(* IEC 61131-3 sources: JingjiangArm/moonboxpro_arm_8.4/Application/Application/任务列表/LogTask/粗采样保存/调用功能, 2 files *)

(* ---- KS_FetchNextSampleDataPtr.st ---- *)
(*@CES
Name=KS_FetchNextSampleDataPtr
Type=FunctionBlock
TypeGuid=6f9dac99-8de1-4efc-8465-68ac443b7d08
Guid=600b6e6a-0af7-4a30-ab9c-796b863be3cd
HasDeclaration=True
HasImplementation=True
*)
{DECLARATION}
FUNCTION KS_FetchNextSampleDataPtr : BOOL
VAR_INPUT
	i_pstStSampleDataForTest: POINTER TO StSampleDataForTest;
	i_ppbyRS_T1: POINTER TO POINTER TO BYTE;(* 粗采样T1数据起点 *)
	i_ppbyRS_T2: POINTER TO POINTER TO BYTE;(* 粗采样T2数据起点 *)
	i_ppbyFS_T1: POINTER TO POINTER TO BYTE;(* 精采样T1数据起点 *)
	i_ppbyFS_T2: POINTER TO POINTER TO BYTE;(* 精采样T2数据起点 *)
END_VAR
VAR
	xResult: BOOL;
	byIDX_Tmp: BYTE;
END_VAR
{IMPLEMENTATION}
IF i_pstStSampleDataForTest<>0 AND
	i_ppbyRS_T1<>0 AND
	i_ppbyRS_T2<>0 AND
	i_ppbyFS_T1<>0 AND
	i_ppbyFS_T2<>0 THEN

	xResult:= TRUE;

	(* 将当前数据位置反馈到出口参数 *)
	byIDX_Tmp:= i_pstStSampleDataForTest^.byIdx AND 7;(* 只取低3位 *)

	(* 粗采样 *)
	i_ppbyRS_T1^:= ADR(i_pstStSampleDataForTest^.abyBuf_Rs[byIDX_Tmp,   1]);
	i_ppbyRS_T2^:= ADR(i_pstStSampleDataForTest^.abyBuf_Rs[byIDX_Tmp,4001]);

	(* 精采样 *)
	i_ppbyFS_T1^:= ADR(i_pstStSampleDataForTest^.abyBuf_Fs[byIDX_Tmp,   1]);
	i_ppbyFS_T2^:= ADR(i_pstStSampleDataForTest^.abyBuf_Fs[byIDX_Tmp,4001]);

	(* go next *)
	i_pstStSampleDataForTest^.byIdx:= i_pstStSampleDataForTest^.byIdx+1;
ELSE
	xResult:= FALSE;
END_IF
KS_FetchNextSampleDataPtr:= xResult;

(* ---- KS_MallocMemAndInstallSampleDataFromFile.st ---- *)
(*@CES
Name=KS_MallocMemAndInstallSampleDataFromFile
Type=FunctionBlock
TypeGuid=6f9dac99-8de1-4efc-8465-68ac443b7d08
Guid=69c33b95-f0e0-43d2-8407-04367f5534f4
HasDeclaration=True
HasImplementation=True
*)
{DECLARATION}
FUNCTION KS_MallocMemAndInstallSampleDataFromFile : DWORD
VAR_INPUT
	i_sFilename_Rs_demo: STRING := '\cpac\rs.demo';
	i_sFilename_Fs_demo: STRING := '\cpac\fs.demo';
END_VAR
VAR
	iN: INT;
	dwMemHdl: DWORD;(* 内存句柄 *)
	dwFileHdl: DWORD;(* 文件句柄 *)
	diSize_Rs_demo: DINT;
	diSize_Fs_demo: DINT;
	pstStSampleDataForTest: POINTER TO StSampleDataForTest := 0;
END_VAR
{IMPLEMENTATION}
dwMemHdl:= SysMemAlloc(SIZEOF(pstStSampleDataForTest^));
pstStSampleDataForTest:= dwMemHdl;
IF pstStSampleDataForTest<>0 THEN
	(* 粗采样 *)
	diSize_Rs_demo:= SysFileGetSize(i_sFilename_Rs_demo);
	IF diSize_Rs_demo=16#10000 THEN(* 文件必须64kB *)
		dwFileHdl:= SysFileOpen(i_sFilename_Rs_demo, 'r');
		IF dwFileHdl<>0 THEN
			FOR iN:=1 TO 8 BY 1 DO
				SysFileSetPos(dwFileHdl, INT_TO_DWORD(iN-1)*8192);(* T1 *)
				SysFileRead(dwFileHdl, ADR(pstStSampleDataForTest^.abyBuf_Rs[iN-1,   1]), 4000);
				SysFileSetPos(dwFileHdl, INT_TO_DWORD(iN-1)*8192+4096);(* T2 *)
				SysFileRead(dwFileHdl, ADR(pstStSampleDataForTest^.abyBuf_Rs[iN-1,4001]), 4000);
			END_FOR
			SysFileClose(dwFileHdl);
		END_IF
	END_IF

	(* 精采样 *)
	diSize_Fs_demo:= SysFileGetSize(i_sFilename_Fs_demo);
	IF diSize_Fs_demo=16#10000 THEN(* 文件必须64kB *)
		dwFileHdl:= SysFileOpen(i_sFilename_Fs_demo, 'r');
		IF dwFileHdl<>0 THEN
			FOR iN:=1 TO 8 BY 1 DO
				SysFileSetPos(dwFileHdl, INT_TO_DWORD(iN-1)*8192);(* T1 *)
				SysFileRead(dwFileHdl, ADR(pstStSampleDataForTest^.abyBuf_Fs[iN-1,   1]), 4000);
				SysFileSetPos(dwFileHdl, INT_TO_DWORD(iN-1)*8192+4096);(* T2 *)
				SysFileRead(dwFileHdl, ADR(pstStSampleDataForTest^.abyBuf_Fs[iN-1,4001]), 4000);
			END_FOR
			SysFileClose(dwFileHdl);
		END_IF
	END_IF
END_IF
KS_MallocMemAndInstallSampleDataFromFile:= dwMemHdl;
